// TIA Portal V20 export
VAR_GLOBAL   // PLC tag table "PLC-A4-DI"
   "-KA6" AT %I8.0 : Bool;
   "-KA7" AT %I8.1 : Bool;
   "-KA8" AT %I8.2 : Bool;
   "-KA9" AT %I8.3 : Bool;
   "-KA10" AT %I8.4 : Bool;
   "-KA11" AT %I8.5 : Bool;
   RESERVE_DI_9 AT %I8.6 : Bool;
   RESERVE_DI_10 AT %I8.7 : Bool;
   RESERVE_DI_11 AT %I9.0 : Bool;   // dveře L kanál A
   RESERVE_DI_12 AT %I9.1 : Bool;   // dveře L kanál B
   RESERVE_DI_13 AT %I9.2 : Bool;   // dveře P kanál A
   RESERVE_DI_14 AT %I9.3 : Bool;   // Dveře P kanál B
   RESERVE_DI_15 AT %I9.4 : Bool;
   RESERVE_DI_16 AT %I9.5 : Bool;
   RESERVE_DI_17 AT %I9.6 : Bool;
   RESERVE_DI_18 AT %I9.7 : Bool;
END_VAR
